ABB RobotStudio station: Prßctica2.rspag

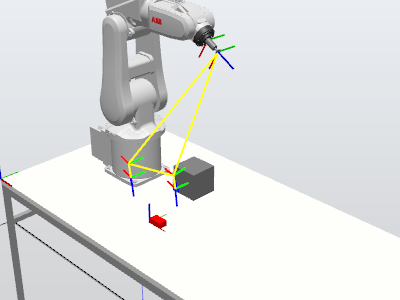
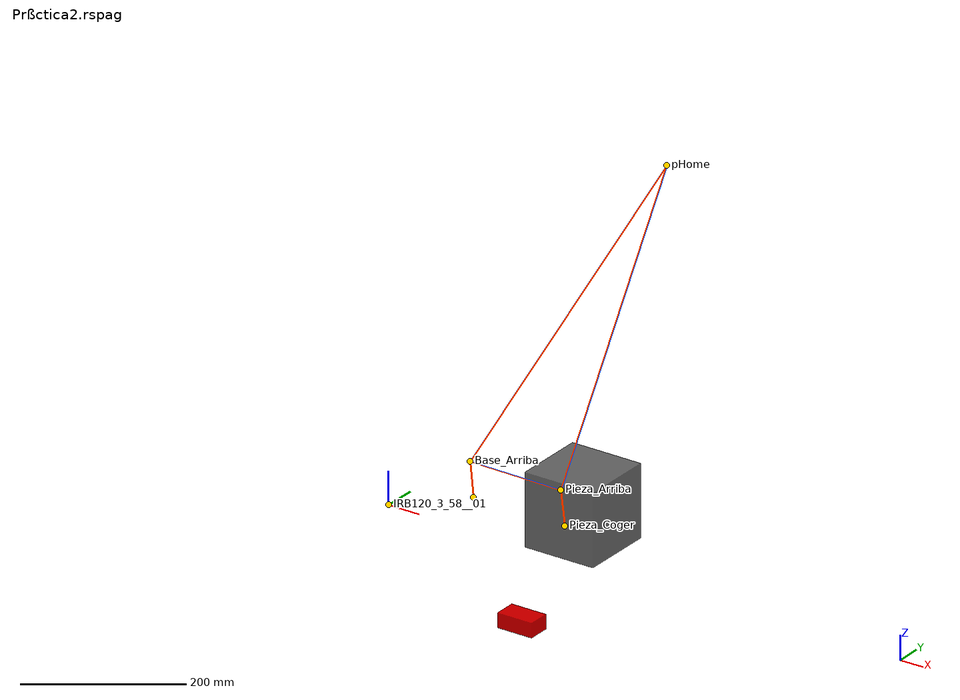
[picture v1: parts stored in the station drawn from their meshes, with robot base, taught points and paths (robot models come from the ABB library and are not in the file)]
--- station ---
Station Práctica2 (saved by RobotStudio 25.4.11475.0)
Controller Controlador2, task T_ROB1: task frame (RAPID world) sits at (0, 0, 670) mm in the station
Controller Controlador2
  mechanical unit ROB_1: IRB120_3_58__01, 6 joints, base frame (0, 0, 0) mm
Layout (positions relative to the parent item):
  - TVentosa [mechanism] at (364.35, 0, 1264) mm, rotated rx 180 ry 60 rz 180 deg
      TCP TVentosa at (0, 0, 51.19) mm
      links: Mi_herramienta
  - LogicGate [smart component, from Components\LogicGate.rslib]
      properties: Operator=NOT; Delay=0
  - LogicGate_2 [smart component, from Components\LogicGate.rslib]
      properties: Operator=AND; Delay=0
  - IRB120_3_58__01 [mechanism, from %ABB.RobotStudio.Models.IRB120%\IRB120_3_58_G_01.rslib] at (0, 0, 670) mm; joint values [0, 0, 0, 0, 0.5236, 0] (rad or m)
  - table [part, from Libraries\Table.rslib] at (-300, 308.26, 670) mm, rotated rx 0 ry 0 rz -90 deg
  - Pieza [part] at (325, -185, 690) mm, rotated rx -180 ry 0 rz 180 deg, size 50 x 30 x 20 mm
  - Base [part], size 100 x 100 x 100 mm
  - Attacher [smart component, from Components\Attacher.rslib]
      properties: Parent=TVentosa; Flange=0; Child=Pieza; Mount=true; Offset=[0 0 0]; Orientation=[0 0 0]
  - CollisionSensor [smart component, from Components\CollisionSensor.rslib]
      properties: Object1=TVentosa; Object2=Pieza; NearMiss=0.001; Part1=(none); Part2=(none); CollisionType=0
    - _sensorPart_ [part]
  - Detacher [smart component, from Components\Detacher.rslib]
      properties: Child=Pieza; KeepPosition=true
Attachment: TVentosa is attached to IRB120_3_58__01 / Link6
Attachment: WO_Base is attached to Base
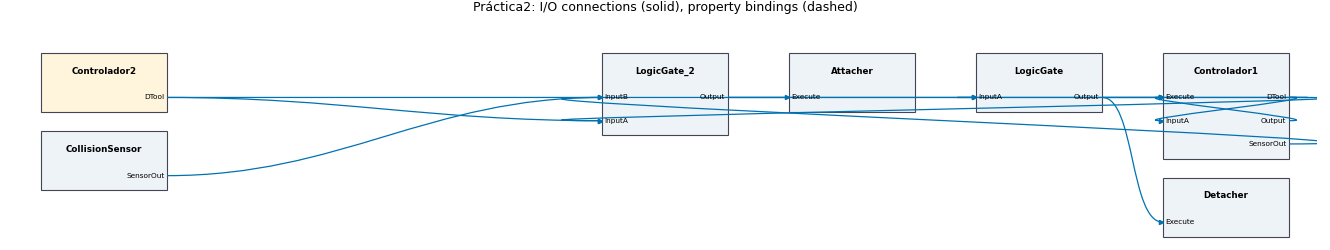
Station logic (signal -> signal, property => property):
  Controlador1.DTool -> Attacher.Execute
  Controlador1.DTool -> LogicGate_2.InputA
  LogicGate_2.Output -> Detacher.Execute
  Controlador1.DTool -> LogicGate.InputA
  LogicGate.Output -> Detacher.Execute
  CollisionSensor.SensorOut -> LogicGate_2.InputB
  Controlador1.DTool -> LogicGate_2.InputA
  LogicGate_2.Output -> Attacher.Execute
  Controlador2.DTool -> LogicGate_2.InputA
  CollisionSensor.SensorOut -> LogicGate_2.InputB
  LogicGate_2.Output -> Attacher.Execute
  LogicGate.Output -> Detacher.Execute
  Controlador2.DTool -> LogicGate.InputA

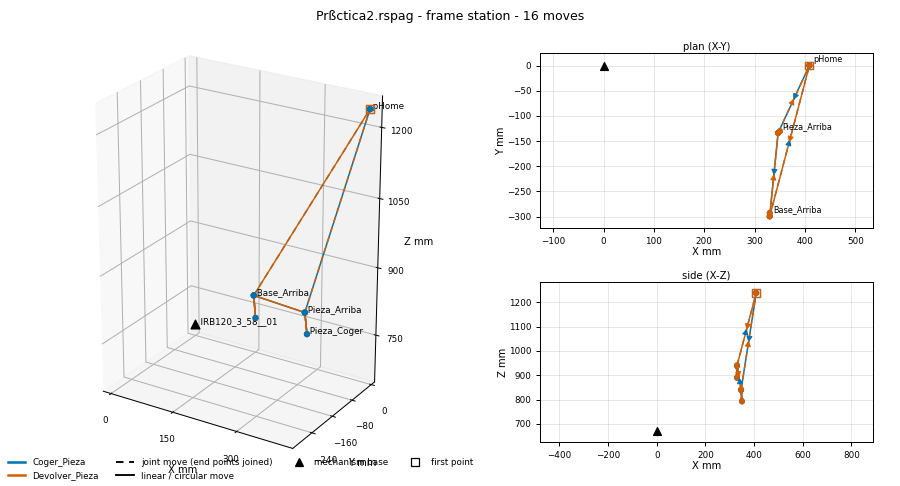
[picture p0: tool path of Prßctica2.rspag in frame station, 16 of 16 moves have a stored position in this frame; points joined in program order, loops and branches not executed]
--- Backups/Controlador2/RAPID/TASK1/PROGMOD/CalibData.mod ---
MODULE CalibData
    PERS tooldata TVentosa:=[TRUE,[[0,0,135],[1,0,0,0]],[0.1,[0,0,1],[1,0,0,0],0,0,0]];
    TASK PERS wobjdata WO_Pieza:=[FALSE,TRUE,"",[[-299.99997408,-391.743024817,0.046553688],[1,-0.000000004,-0.000000007,0]],[[600,191.743,0],[1,0,0,0]]];
    TASK PERS wobjdata WO_Base:=[FALSE,TRUE,"",[[-300,-391.743,0],[1,0,0,0]],[[500,391.743,0],[1,0,0,0]]];
ENDMODULE

--- Backups/Controlador2/RAPID/TASK1/PROGMOD/Module1.mod ---
MODULE Module1
    CONST robtarget pHome:=[[408.686,0,568.405],[0.5,0,0.866025404,0],[0,0,0,0],[9E+09,9E+09,9E+09,9E+09,9E+09,9E+09]];
    CONST robtarget Pieza_Arriba:=[[46.55,66.15,170.37],[0.030252817,-0.082767664,-0.983572083,-0.157544399],[-1,0,-1,0],[9E+09,9E+09,9E+09,9E+09,9E+09,9E+09]];
    CONST robtarget Pieza_Coger:=[[50.14,69.58,122.36],[0.040345362,-0.101949598,-0.991439425,-0.070897089],[0,0,0,0],[9E+09,9E+09,9E+09,9E+09,9E+09,9E+09]];
    CONST robtarget Base_Arriba:=[[129.83,-299.55,269.95],[0.040354259,-0.101946077,-0.991445608,-0.07081057],[0,0,-2,0],[9E+09,9E+09,9E+09,9E+09,9E+09,9E+09]];
    CONST robtarget Base_Coger:=[[129.88,-292.83,219.57],[0.040267684,-0.101940713,-0.991450276,-0.070802219],[0,0,-2,0],[9E+09,9E+09,9E+09,9E+09,9E+09,9E+09]];

    PROC main()
        Coger_Pieza;
        Devolver_Pieza;
    ENDPROC

    PROC Coger_Pieza()
        MoveJ pHome,v150,fine,TVentosa\WObj:=wobj0;

        MoveL Pieza_Arriba,v150,fine,TVentosa\WObj:=WO_Pieza;
        MoveL Pieza_Coger,v150,fine,TVentosa\WObj:=WO_Pieza;

        WaitTime 0.5;
        SetDO DTool,1;
        WaitTime 0.5;

        MoveL Pieza_Arriba,v150,fine,TVentosa\WObj:=WO_Pieza;
        MoveL Base_Arriba,v150,fine,TVentosa\WObj:=WO_Base;
        MoveL Base_Coger,v150,fine,TVentosa\WObj:=WO_Base;
        WaitTime 0.5;
        SetDO DTool,0;
        WaitTime 0.5;

        MoveL Base_Arriba,v150,fine,TVentosa\WObj:=WO_Base;
        MoveJ pHome,v150,fine,TVentosa\WObj:=wobj0;
    ENDPROC

    PROC Devolver_Pieza()
        MoveJ pHome,v150,fine,TVentosa\WObj:=wobj0;

        MoveL Base_Arriba,v150,fine,TVentosa\WObj:=WO_Base;
        MoveL Base_Coger,v150,fine,TVentosa\WObj:=WO_Base;
        WaitTime 0.5;
        SetDO DTool,1;
        WaitTime 0.5;

        MoveL Base_Arriba,v150,fine,TVentosa\WObj:=WO_Base;
        MoveL Pieza_Arriba,v150,fine,TVentosa\WObj:=WO_Pieza;
        MoveL Pieza_Coger,v150,fine,TVentosa\WObj:=WO_Pieza;

        WaitTime 0.5;
        SetDO DTool,0;
        WaitTime 0.5;
        MoveL Pieza_Arriba,v150,fine,TVentosa\WObj:=WO_Pieza;
        MoveJ pHome,v150,fine,TVentosa\WObj:=wobj0;
    ENDPROC
ENDMODULE

--- Backups/Controlador2/SYSPAR/EIO.cfg ---
EIO:CFG_1.0:6:1::
#
EIO_SIGNAL:

      -Name "DTool" -SignalType "DO"

      -Name "DI0" -SignalType "DI"
